FUNCTION_BLOCK StructProducer
  (* Standard: 61499-1 *)
  (* Version 1.0, 2026-05-26, Dimitrios Kalligaridis *)
  PACKAGE mypackage;
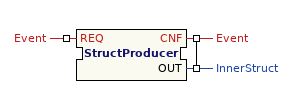
  EVENT_INPUT
    REQ WITH OUT;
  END_EVENT
  EVENT_OUTPUT
    CNF WITH OUT;
  END_EVENT
  VAR_OUTPUT
    OUT : mypackage::InnerStruct;
  END_VAR
  EC_STATES
    START;
  END_STATES
END_FUNCTION_BLOCK
